# EPICS autosave request: iocs/ad/pylon-ioc/db/ADGenICam_settings.req
file "ADBase_settings.req", P=$(P), R=$(R)
$(P)$(R)FrameRateEnable
$(P)$(R)TriggerSource
$(P)$(R)TriggerOverlap
$(P)$(R)ExposureMode
$(P)$(R)ExposureAuto
$(P)$(R)GainAuto
$(P)$(R)PixelFormat
